Fanuc KAREL source: KA00116.KL

PROGRAM KA00116
%NOLOCKGROUP
VAR
  SRC: CONFIG
  DST: JOINTPOS
BEGIN
  SRC.CFG_FLIP = TRUE
  DST = SRC
END KA00116
